// TIA Portal V20 export
DATA_BLOCK "MCP_RC_DB5"   // DB9808
{ S7_Optimized_Access := 'TRUE' }
   VAR
      Count : Int := 5;
      D : "MCP_RC_UDTD";
   END_VAR
BEGIN
END_DATA_BLOCK
